SUBAPPLICATION AE_AX_SERVER_0_PUBLISH_1 (* Wie adapter::net::AE_AX_SERVER_0_CLIENT_1_0, aber lokales PUBLISH_1 statt Remote-CLIENT_1_0 (ein Geraet) *)
  (* Standard: 61499-2; Description: Copyright (c) 2026 HR Agrartechnik GmbH This program and the accompanying materials are made available under the terms of the Eclipse Public License 2.0 which is available at https://www.eclipse.org/legal/epl-2.0/ SPDX-License-Identifier: EPL-2.0 *)
  (* Version 1.2, 2026-11-25, Franz Höpfinger, Meisterschulen am Ostbahnhof, SERVER_0 -> MyLib::net::SERVER_0_QO (IND nur bei QO=TRUE, RSP intern). Ein gescheitertes RSP meldet IND mit QO=FALSE, direkt IND->RSP ergab eine Endlosschleife. *)
  (* Version 1.1, 2026-10-18, Franz Höpfinger, Meisterschulen am Ostbahnhof, Kopie von AE_AX_SERVER_0_CLIENT_1_0, CLIENT_1_0 durch PUBLISH_1 ersetzt - als SubAppType, damit FORTE den Typ nicht kennen muss (kein ELF fuer MyLib_AX). SERVER_0: IND direkt auf RSP (sonst bis 4 s Server-Lock fuer alle Publishes) *)
  (* Version 1.0, 2026-09-03, Franz Höpfinger, HR Agrartechnik GmbH, initial API and implementation and/or initial documentation *)
  PACKAGE MyLib::net;
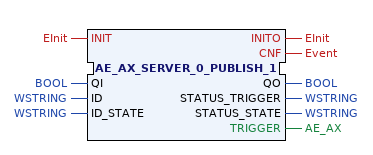
  EVENT_INPUT
    INIT : EInit; (* Initialization *)
  END_EVENT
  EVENT_OUTPUT
    INITO : EInit; (* Initialization Confirm *)
    CNF; (* QO/STATUS updated *)
  END_EVENT
  VAR_INPUT
    QI : BOOL;
    ID : WSTRING; (* Lokale Methodenadresse (ACTION=CREATE_METHOD) fuer den Trigger-Methodenaufruf *)
    ID_STATE : WSTRING; (* Lokale Adresse (ACTION=WRITE) fuer den Zustand *)
  END_VAR
  VAR_OUTPUT
    QO : BOOL; (* TRUE nur wenn SERVER_0_1 und STATE_CLIENT aktuell beide QO=TRUE melden *)
    STATUS_TRIGGER : WSTRING; (* STATUS von SERVER_0_1 *)
    STATUS_STATE : WSTRING; (* STATUS von STATE_CLIENT *)
  END_VAR
  PLUGS
    TRIGGER : adapter::types::bidirectional::AE_AX; (* Trigger (in), Zustand (out) *)
  END_PLUGS
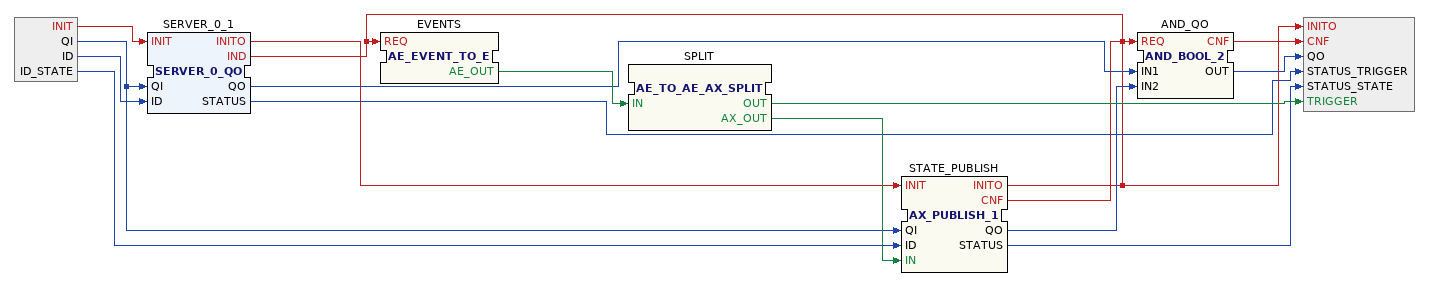
  FBS
    EVENTS : adapter::conversion::unidirectional::AE_EVENT_TO_E;
    SPLIT : adapter::events::bidirectional::AE_TO_AE_AX_SPLIT;
    STATE_PUBLISH : adapter::net::AX_PUBLISH_1;
    AND_QO : iec61131::booleanOperators::AND_BOOL_2;
  END_FBS
  SUBAPPS
    SERVER_0_1 : MyLib::net::SERVER_0_QO;
  END_SUBAPPS
  EVENT_CONNECTIONS
    INIT TO SERVER_0_1.INIT;
    SERVER_0_1.INITO TO STATE_PUBLISH.INIT;
    STATE_PUBLISH.INITO TO INITO;
    STATE_PUBLISH.INITO TO AND_QO.REQ;
    SERVER_0_1.IND TO EVENTS.REQ;
    SERVER_0_1.IND TO AND_QO.REQ;
    STATE_PUBLISH.CNF TO AND_QO.REQ;
    AND_QO.CNF TO CNF;
  END_CONNECTIONS
  DATA_CONNECTIONS
    QI TO SERVER_0_1.QI;
    ID TO SERVER_0_1.ID;
    SERVER_0_1.QO TO AND_QO.IN1;
    SERVER_0_1.STATUS TO STATUS_TRIGGER;
    QI TO STATE_PUBLISH.QI;
    ID_STATE TO STATE_PUBLISH.ID;
    STATE_PUBLISH.QO TO AND_QO.IN2;
    AND_QO.OUT TO QO;
    STATE_PUBLISH.STATUS TO STATUS_STATE;
  END_CONNECTIONS
  ADAPTER_CONNECTIONS
    EVENTS.AE_OUT TO SPLIT.IN;
    SPLIT.OUT TO TRIGGER;
    SPLIT.AX_OUT TO STATE_PUBLISH.IN;
  END_CONNECTIONS
END_SUBAPPLICATION
